Fanuc KAREL source: kd00048.KL

-- PROVISIONAL review KL for V770-1; original PC SHA256 1dd4873eb4a397bb0ae44bab8086c2c37b592e7663dd33b537e2391eae96038e
-- Incomplete behavior may be omitted. Consult companion uncertainty JSON. Do not deploy.
PROGRAM KD00048
%NOLOCKGROUP
BEGIN
  -- UNRESOLVED_PC offsets 5-29; opcodes 01,22,1C,9D,2C,08,82,0B
  -- UNRESOLVED_PC offsets 34-38; opcodes 7F
END KD00048
